// TIA Portal V20 export
FUNCTION_BLOCK "PR_FibroMainSeq_Soft2.0 1_workflow_a30ae2"   // FB43, LAD
{ S7_Optimized_Access := 'TRUE' }
// stored: MemoryReserve 100, SetENOAutomatically false
   VAR_INPUT
      iAllStationsSafe : Bool;
      iAllTaskOver : Bool;
      iAutoRunning : Bool;
      iFaultReset : Bool;
      iFibroAtStnPos : Bool;
      iIndexOver : Bool;
      iProcessActive : Bool;
      iReset_fault : Bool;
      iSstMode : Bool;
      iSstPB : Bool;
   END_VAR
   VAR_OUTPUT
      qError : Array[1..1] of Bool;
      qMessage_0 : Bool;
      qProcessActive : Bool;
   END_VAR
   VAR
      c10_ChkRecCond_T1 : Bool;
      c10_ChkRecCond_T2 : Bool;
      c10_ChkRecCond_T3 : Bool;
      c50_ChkPartPresentAtStn_T1 : Bool;
      c50_ChkPartPresentAtStn_T2 : Bool;
      StateNo : Int;
      s100_WtAllStnTaskOver : Bool;
      s100_WtAllStnTaskOver_T1 : Bool;
      s10_ChkRecCond : Bool;
      s10_ChkRecCond_T1 : Bool;
      s10_ChkRecCond_T2 : Bool;
      s10_ChkRecCond_T3 : Bool;
      s130_ChkAllStnSafe2 : Bool;
      s130_ChkAllStnSafe2_T1 : Bool;
      s140_WtIndexOver : Bool;
      s140_WtIndexOver_T1 : Bool;
      s1_WtResetRel : Bool;
      s1_WtResetRel_T1 : Bool;
      s20_WtManualIntv : Bool;
      s20_WtManualIntv_T1 : Bool;
      s30_WtFibroAtStnPos : Bool;
      s30_WtFibroAtStnPos_T1 : Bool;
      s40_ChkAllStnSafe : Bool;
      s40_ChkAllStnSafe_T1 : Bool;
      s50_ChkPartPresentAtStn : Bool;
      s50_ChkPartPresentAtStn_T1 : Bool;
      s50_ChkPartPresentAtStn_T2 : Bool;
      s60_WtPartPresentAtStn : Bool;
      s60_WtPartPresentAtStn_T1 : Bool;
      sAbnormalCondition : Bool;
      sPartPresentAtStation : Bool;
      sProcessActive : Bool;
      sSst : Bool;
      sSstPulse : Bool;
      sSstRise : Bool;
      sStWtResetRel : Bool;
      sStWtResetRel_T1 : Bool;
   END_VAR
   VAR_TEMP
      tOne : Bool;
   END_VAR
   VAR_TEMP   // added for the SCL form of the ladder/FBD networks
      _w1 : Bool;
      _w2 : Bool;
   END_VAR
BEGIN

REGION Network 1
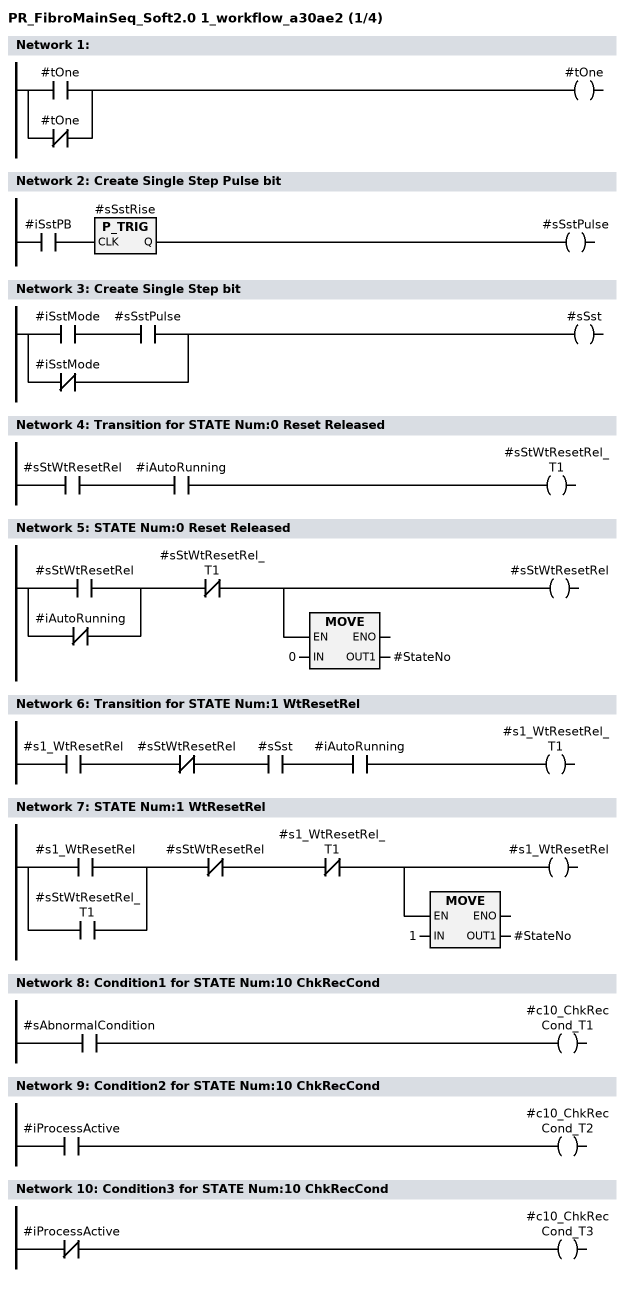
   RUNG wire#powerrail
      Contact( #tOne )
      wire#w1
      Coil( #tOne )
   END_RUNG
   RUNG wire#powerrail
      I_Contact( #tOne )
   END_RUNG wire#w1
   // the same network as SCL:
   #tOne := #tOne OR NOT #tOne;
END_REGION

REGION Network 2: Create Single Step Pulse bit
   RUNG wire#powerrail
      Contact( #iSstPB )
      P_Trig( #sSstRise )
      Coil( #sSstPulse )
   END_RUNG
   // the same network as SCL:
   #_w1 := #iSstPB AND NOT #sSstRise;   // rising edge
   #sSstRise := #iSstPB;
   #sSstPulse := #_w1;
END_REGION

REGION Network 3: Create Single Step bit
   RUNG wire#powerrail
      Contact( #iSstMode )
      Contact( #sSstPulse )
      wire#w1
      Coil( #sSst )
   END_RUNG
   RUNG wire#powerrail
      I_Contact( #iSstMode )
   END_RUNG wire#w1
   // the same network as SCL:
   #sSst := (#iSstMode AND #sSstPulse) OR NOT #iSstMode;
END_REGION

REGION Network 4: Transition for STATE Num:0 Reset Released
   RUNG wire#powerrail
      Contact( #sStWtResetRel )
      Contact( #iAutoRunning )
      Coil( #sStWtResetRel_T1 )
   END_RUNG
   // the same network as SCL:
   #sStWtResetRel_T1 := #sStWtResetRel AND #iAutoRunning;
END_REGION

REGION Network 5: STATE Num:0 Reset Released
   RUNG wire#powerrail
      Contact( #sStWtResetRel )
      wire#w1
      I_Contact( #sStWtResetRel_T1 )
      wire#w2
      Coil( #sStWtResetRel )
   END_RUNG
   RUNG wire#powerrail
      I_Contact( #iAutoRunning )
   END_RUNG wire#w1
   RUNG wire#w2
      { S7_GenerateENO := "TRUE" } Move(in := 0, out1 => #StateNo)
   END_RUNG
   // the same network as SCL:
   #sStWtResetRel := (#sStWtResetRel OR NOT #iAutoRunning) AND NOT #sStWtResetRel_T1;
   IF #sStWtResetRel THEN #StateNo := 0; END_IF;
END_REGION

REGION Network 6: Transition for STATE Num:1 WtResetRel
   RUNG wire#powerrail
      Contact( #s1_WtResetRel )
      I_Contact( #sStWtResetRel )
      Contact( #sSst )
      Contact( #iAutoRunning )
      Coil( #s1_WtResetRel_T1 )
   END_RUNG
   // the same network as SCL:
   #s1_WtResetRel_T1 := #s1_WtResetRel AND NOT #sStWtResetRel AND #sSst AND #iAutoRunning;
END_REGION

REGION Network 7: STATE Num:1 WtResetRel
   RUNG wire#powerrail
      Contact( #s1_WtResetRel )
      wire#w1
      I_Contact( #sStWtResetRel )
      I_Contact( #s1_WtResetRel_T1 )
      wire#w2
      Coil( #s1_WtResetRel )
   END_RUNG
   RUNG wire#powerrail
      Contact( #sStWtResetRel_T1 )
   END_RUNG wire#w1
   RUNG wire#w2
      { S7_GenerateENO := "TRUE" } Move(in := 1, out1 => #StateNo)
   END_RUNG
   // the same network as SCL:
   #s1_WtResetRel := (#s1_WtResetRel OR #sStWtResetRel_T1) AND NOT #sStWtResetRel AND NOT #s1_WtResetRel_T1;
   IF #s1_WtResetRel THEN #StateNo := 1; END_IF;
END_REGION

REGION Network 8: Condition1 for STATE Num:10 ChkRecCond
   RUNG wire#powerrail
      Contact( #sAbnormalCondition )
      Coil( #c10_ChkRecCond_T1 )
   END_RUNG
   // the same network as SCL:
   #c10_ChkRecCond_T1 := #sAbnormalCondition;
END_REGION

REGION Network 9: Condition2 for STATE Num:10 ChkRecCond
   RUNG wire#powerrail
      Contact( #iProcessActive )
      Coil( #c10_ChkRecCond_T2 )
   END_RUNG
   // the same network as SCL:
   #c10_ChkRecCond_T2 := #iProcessActive;
END_REGION

REGION Network 10: Condition3 for STATE Num:10 ChkRecCond
   RUNG wire#powerrail
      I_Contact( #iProcessActive )
      Coil( #c10_ChkRecCond_T3 )
   END_RUNG
   // the same network as SCL:
   #c10_ChkRecCond_T3 := NOT #iProcessActive;
END_REGION

REGION Network 11: Transition for STATE Num:10 ChkRecCond
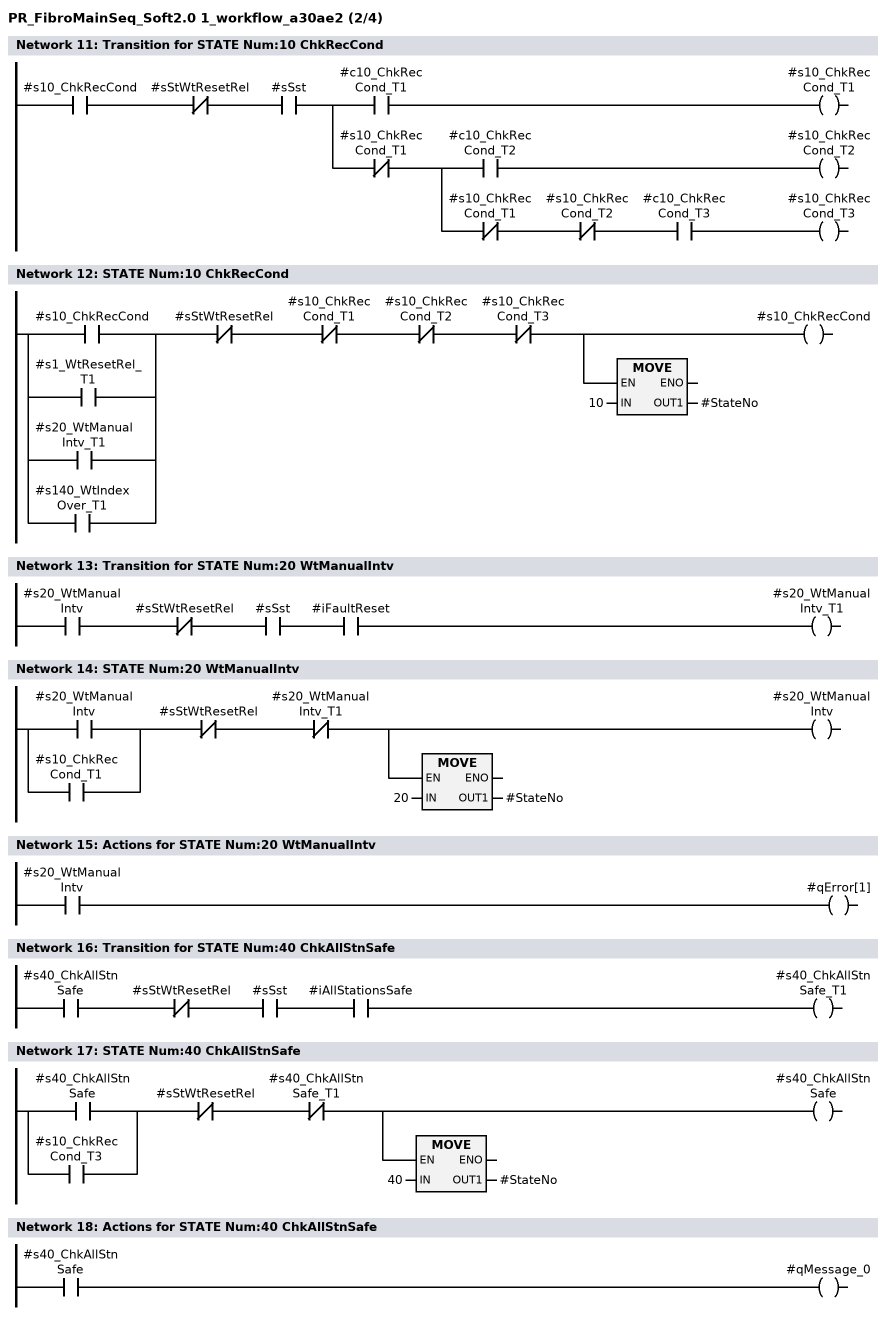
   RUNG wire#powerrail
      Contact( #s10_ChkRecCond )
      I_Contact( #sStWtResetRel )
      Contact( #sSst )
      wire#w1
      Contact( #c10_ChkRecCond_T1 )
      Coil( #s10_ChkRecCond_T1 )
   END_RUNG
   RUNG wire#w1
      I_Contact( #s10_ChkRecCond_T1 )
      wire#w2
      Contact( #c10_ChkRecCond_T2 )
      Coil( #s10_ChkRecCond_T2 )
   END_RUNG
   RUNG wire#w2
      I_Contact( #s10_ChkRecCond_T1 )
      I_Contact( #s10_ChkRecCond_T2 )
      Contact( #c10_ChkRecCond_T3 )
      Coil( #s10_ChkRecCond_T3 )
   END_RUNG
   // the same network as SCL:
   #_w1 := #s10_ChkRecCond AND NOT #sStWtResetRel AND #sSst;
   #s10_ChkRecCond_T1 := #_w1 AND #c10_ChkRecCond_T1;
   #_w2 := #_w1 AND NOT #s10_ChkRecCond_T1;
   #s10_ChkRecCond_T2 := #_w2 AND #c10_ChkRecCond_T2;
   #s10_ChkRecCond_T3 := #_w2 AND NOT #s10_ChkRecCond_T1 AND NOT #s10_ChkRecCond_T2 AND #c10_ChkRecCond_T3;
END_REGION

REGION Network 12: STATE Num:10 ChkRecCond
   RUNG wire#powerrail
      Contact( #s10_ChkRecCond )
      wire#w1
      I_Contact( #sStWtResetRel )
      I_Contact( #s10_ChkRecCond_T1 )
      I_Contact( #s10_ChkRecCond_T2 )
      I_Contact( #s10_ChkRecCond_T3 )
      wire#w2
      Coil( #s10_ChkRecCond )
   END_RUNG
   RUNG wire#powerrail
      Contact( #s1_WtResetRel_T1 )
   END_RUNG wire#w1
   RUNG wire#powerrail
      Contact( #s20_WtManualIntv_T1 )
   END_RUNG wire#w1
   RUNG wire#powerrail
      Contact( #s140_WtIndexOver_T1 )
   END_RUNG wire#w1
   RUNG wire#w2
      { S7_GenerateENO := "TRUE" } Move(in := 10, out1 => #StateNo)
   END_RUNG
   // the same network as SCL:
   #s10_ChkRecCond := (#s10_ChkRecCond OR #s1_WtResetRel_T1 OR #s20_WtManualIntv_T1 OR #s140_WtIndexOver_T1) AND NOT #sStWtResetRel AND NOT #s10_ChkRecCond_T1 AND NOT #s10_ChkRecCond_T2 AND NOT #s10_ChkRecCond_T3;
   IF #s10_ChkRecCond THEN #StateNo := 10; END_IF;
END_REGION

REGION Network 13: Transition for STATE Num:20 WtManualIntv
   RUNG wire#powerrail
      Contact( #s20_WtManualIntv )
      I_Contact( #sStWtResetRel )
      Contact( #sSst )
      Contact( #iFaultReset )
      Coil( #s20_WtManualIntv_T1 )
   END_RUNG
   // the same network as SCL:
   #s20_WtManualIntv_T1 := #s20_WtManualIntv AND NOT #sStWtResetRel AND #sSst AND #iFaultReset;
END_REGION

REGION Network 14: STATE Num:20 WtManualIntv
   RUNG wire#powerrail
      Contact( #s20_WtManualIntv )
      wire#w1
      I_Contact( #sStWtResetRel )
      I_Contact( #s20_WtManualIntv_T1 )
      wire#w2
      Coil( #s20_WtManualIntv )
   END_RUNG
   RUNG wire#powerrail
      Contact( #s10_ChkRecCond_T1 )
   END_RUNG wire#w1
   RUNG wire#w2
      { S7_GenerateENO := "TRUE" } Move(in := 20, out1 => #StateNo)
   END_RUNG
   // the same network as SCL:
   #s20_WtManualIntv := (#s20_WtManualIntv OR #s10_ChkRecCond_T1) AND NOT #sStWtResetRel AND NOT #s20_WtManualIntv_T1;
   IF #s20_WtManualIntv THEN #StateNo := 20; END_IF;
END_REGION

REGION Network 15: Actions for STATE Num:20 WtManualIntv
   RUNG wire#powerrail
      Contact( #s20_WtManualIntv )
      Coil( #qError[1] )
   END_RUNG
   // the same network as SCL:
   #qError[1] := #s20_WtManualIntv;
END_REGION

REGION Network 16: Transition for STATE Num:40 ChkAllStnSafe
   RUNG wire#powerrail
      Contact( #s40_ChkAllStnSafe )
      I_Contact( #sStWtResetRel )
      Contact( #sSst )
      Contact( #iAllStationsSafe )
      Coil( #s40_ChkAllStnSafe_T1 )
   END_RUNG
   // the same network as SCL:
   #s40_ChkAllStnSafe_T1 := #s40_ChkAllStnSafe AND NOT #sStWtResetRel AND #sSst AND #iAllStationsSafe;
END_REGION

REGION Network 17: STATE Num:40 ChkAllStnSafe
   RUNG wire#powerrail
      Contact( #s40_ChkAllStnSafe )
      wire#w1
      I_Contact( #sStWtResetRel )
      I_Contact( #s40_ChkAllStnSafe_T1 )
      wire#w2
      Coil( #s40_ChkAllStnSafe )
   END_RUNG
   RUNG wire#powerrail
      Contact( #s10_ChkRecCond_T3 )
   END_RUNG wire#w1
   RUNG wire#w2
      { S7_GenerateENO := "TRUE" } Move(in := 40, out1 => #StateNo)
   END_RUNG
   // the same network as SCL:
   #s40_ChkAllStnSafe := (#s40_ChkAllStnSafe OR #s10_ChkRecCond_T3) AND NOT #sStWtResetRel AND NOT #s40_ChkAllStnSafe_T1;
   IF #s40_ChkAllStnSafe THEN #StateNo := 40; END_IF;
END_REGION

REGION Network 18: Actions for STATE Num:40 ChkAllStnSafe
   RUNG wire#powerrail
      Contact( #s40_ChkAllStnSafe )
      Coil( #qMessage_0 )
   END_RUNG
   // the same network as SCL:
   #qMessage_0 := #s40_ChkAllStnSafe;
END_REGION

REGION Network 19: Transition for STATE Num:30 WtFibroAtStnPos
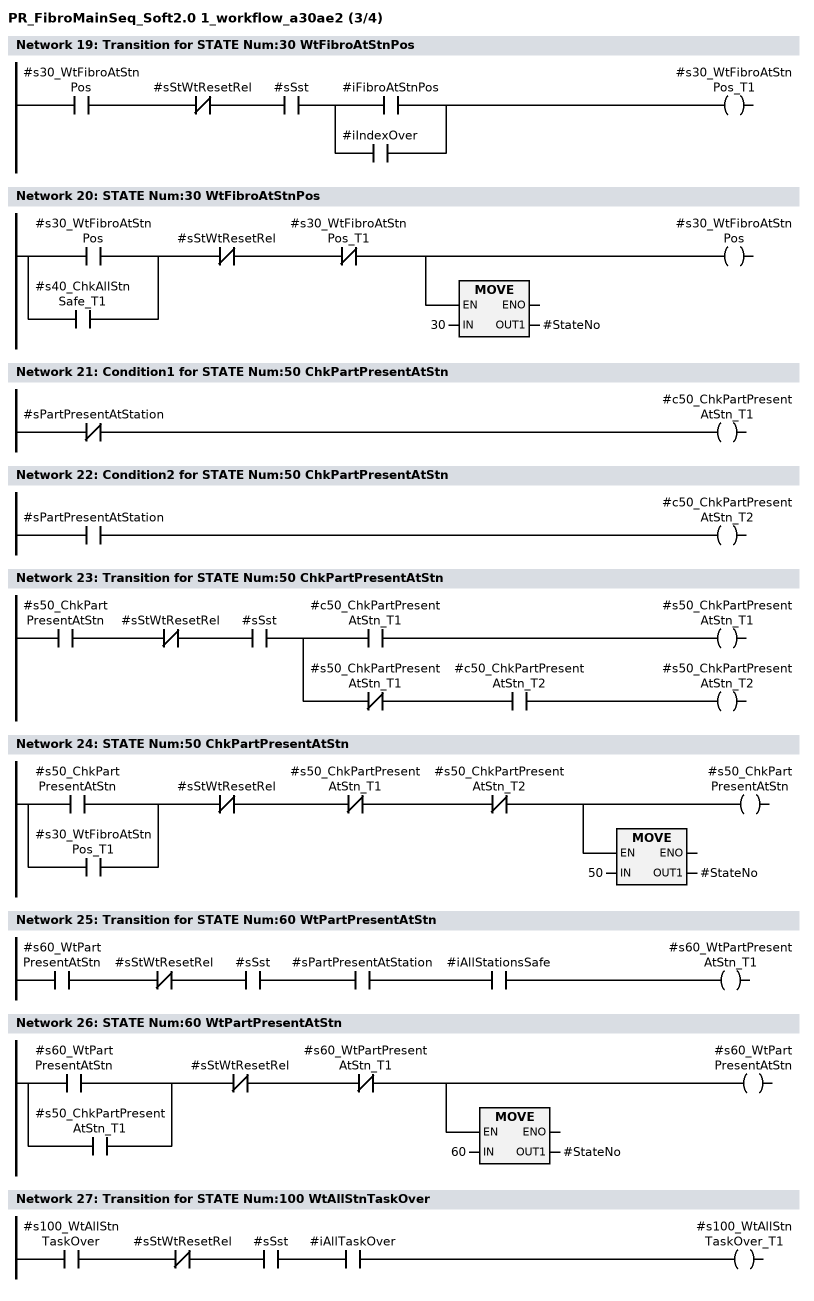
   RUNG wire#powerrail
      Contact( #s30_WtFibroAtStnPos )
      I_Contact( #sStWtResetRel )
      Contact( #sSst )
      wire#w1
      Contact( #iFibroAtStnPos )
      wire#w2
      Coil( #s30_WtFibroAtStnPos_T1 )
   END_RUNG
   RUNG wire#w1
      Contact( #iIndexOver )
   END_RUNG wire#w2
   // the same network as SCL:
   #s30_WtFibroAtStnPos_T1 := #s30_WtFibroAtStnPos AND NOT #sStWtResetRel AND #sSst AND (#iFibroAtStnPos OR #iIndexOver);
END_REGION

REGION Network 20: STATE Num:30 WtFibroAtStnPos
   RUNG wire#powerrail
      Contact( #s30_WtFibroAtStnPos )
      wire#w1
      I_Contact( #sStWtResetRel )
      I_Contact( #s30_WtFibroAtStnPos_T1 )
      wire#w2
      Coil( #s30_WtFibroAtStnPos )
   END_RUNG
   RUNG wire#powerrail
      Contact( #s40_ChkAllStnSafe_T1 )
   END_RUNG wire#w1
   RUNG wire#w2
      { S7_GenerateENO := "TRUE" } Move(in := 30, out1 => #StateNo)
   END_RUNG
   // the same network as SCL:
   #s30_WtFibroAtStnPos := (#s30_WtFibroAtStnPos OR #s40_ChkAllStnSafe_T1) AND NOT #sStWtResetRel AND NOT #s30_WtFibroAtStnPos_T1;
   IF #s30_WtFibroAtStnPos THEN #StateNo := 30; END_IF;
END_REGION

REGION Network 21: Condition1 for STATE Num:50 ChkPartPresentAtStn
   RUNG wire#powerrail
      I_Contact( #sPartPresentAtStation )
      Coil( #c50_ChkPartPresentAtStn_T1 )
   END_RUNG
   // the same network as SCL:
   #c50_ChkPartPresentAtStn_T1 := NOT #sPartPresentAtStation;
END_REGION

REGION Network 22: Condition2 for STATE Num:50 ChkPartPresentAtStn
   RUNG wire#powerrail
      Contact( #sPartPresentAtStation )
      Coil( #c50_ChkPartPresentAtStn_T2 )
   END_RUNG
   // the same network as SCL:
   #c50_ChkPartPresentAtStn_T2 := #sPartPresentAtStation;
END_REGION

REGION Network 23: Transition for STATE Num:50 ChkPartPresentAtStn
   RUNG wire#powerrail
      Contact( #s50_ChkPartPresentAtStn )
      I_Contact( #sStWtResetRel )
      Contact( #sSst )
      wire#w1
      Contact( #c50_ChkPartPresentAtStn_T1 )
      Coil( #s50_ChkPartPresentAtStn_T1 )
   END_RUNG
   RUNG wire#w1
      I_Contact( #s50_ChkPartPresentAtStn_T1 )
      Contact( #c50_ChkPartPresentAtStn_T2 )
      Coil( #s50_ChkPartPresentAtStn_T2 )
   END_RUNG
   // the same network as SCL:
   #_w1 := #s50_ChkPartPresentAtStn AND NOT #sStWtResetRel AND #sSst;
   #s50_ChkPartPresentAtStn_T1 := #_w1 AND #c50_ChkPartPresentAtStn_T1;
   #s50_ChkPartPresentAtStn_T2 := #_w1 AND NOT #s50_ChkPartPresentAtStn_T1 AND #c50_ChkPartPresentAtStn_T2;
END_REGION

REGION Network 24: STATE Num:50 ChkPartPresentAtStn
   RUNG wire#powerrail
      Contact( #s50_ChkPartPresentAtStn )
      wire#w1
      I_Contact( #sStWtResetRel )
      I_Contact( #s50_ChkPartPresentAtStn_T1 )
      I_Contact( #s50_ChkPartPresentAtStn_T2 )
      wire#w2
      Coil( #s50_ChkPartPresentAtStn )
   END_RUNG
   RUNG wire#powerrail
      Contact( #s30_WtFibroAtStnPos_T1 )
   END_RUNG wire#w1
   RUNG wire#w2
      { S7_GenerateENO := "TRUE" } Move(in := 50, out1 => #StateNo)
   END_RUNG
   // the same network as SCL:
   #s50_ChkPartPresentAtStn := (#s50_ChkPartPresentAtStn OR #s30_WtFibroAtStnPos_T1) AND NOT #sStWtResetRel AND NOT #s50_ChkPartPresentAtStn_T1 AND NOT #s50_ChkPartPresentAtStn_T2;
   IF #s50_ChkPartPresentAtStn THEN #StateNo := 50; END_IF;
END_REGION

REGION Network 25: Transition for STATE Num:60 WtPartPresentAtStn
   RUNG wire#powerrail
      Contact( #s60_WtPartPresentAtStn )
      I_Contact( #sStWtResetRel )
      Contact( #sSst )
      Contact( #sPartPresentAtStation )
      Contact( #iAllStationsSafe )
      Coil( #s60_WtPartPresentAtStn_T1 )
   END_RUNG
   // the same network as SCL:
   #s60_WtPartPresentAtStn_T1 := #s60_WtPartPresentAtStn AND NOT #sStWtResetRel AND #sSst AND #sPartPresentAtStation AND #iAllStationsSafe;
END_REGION

REGION Network 26: STATE Num:60 WtPartPresentAtStn
   RUNG wire#powerrail
      Contact( #s60_WtPartPresentAtStn )
      wire#w1
      I_Contact( #sStWtResetRel )
      I_Contact( #s60_WtPartPresentAtStn_T1 )
      wire#w2
      Coil( #s60_WtPartPresentAtStn )
   END_RUNG
   RUNG wire#powerrail
      Contact( #s50_ChkPartPresentAtStn_T1 )
   END_RUNG wire#w1
   RUNG wire#w2
      { S7_GenerateENO := "TRUE" } Move(in := 60, out1 => #StateNo)
   END_RUNG
   // the same network as SCL:
   #s60_WtPartPresentAtStn := (#s60_WtPartPresentAtStn OR #s50_ChkPartPresentAtStn_T1) AND NOT #sStWtResetRel AND NOT #s60_WtPartPresentAtStn_T1;
   IF #s60_WtPartPresentAtStn THEN #StateNo := 60; END_IF;
END_REGION

REGION Network 27: Transition for STATE Num:100 WtAllStnTaskOver
   RUNG wire#powerrail
      Contact( #s100_WtAllStnTaskOver )
      I_Contact( #sStWtResetRel )
      Contact( #sSst )
      Contact( #iAllTaskOver )
      Coil( #s100_WtAllStnTaskOver_T1 )
   END_RUNG
   // the same network as SCL:
   #s100_WtAllStnTaskOver_T1 := #s100_WtAllStnTaskOver AND NOT #sStWtResetRel AND #sSst AND #iAllTaskOver;
END_REGION

REGION Network 28: STATE Num:100 WtAllStnTaskOver
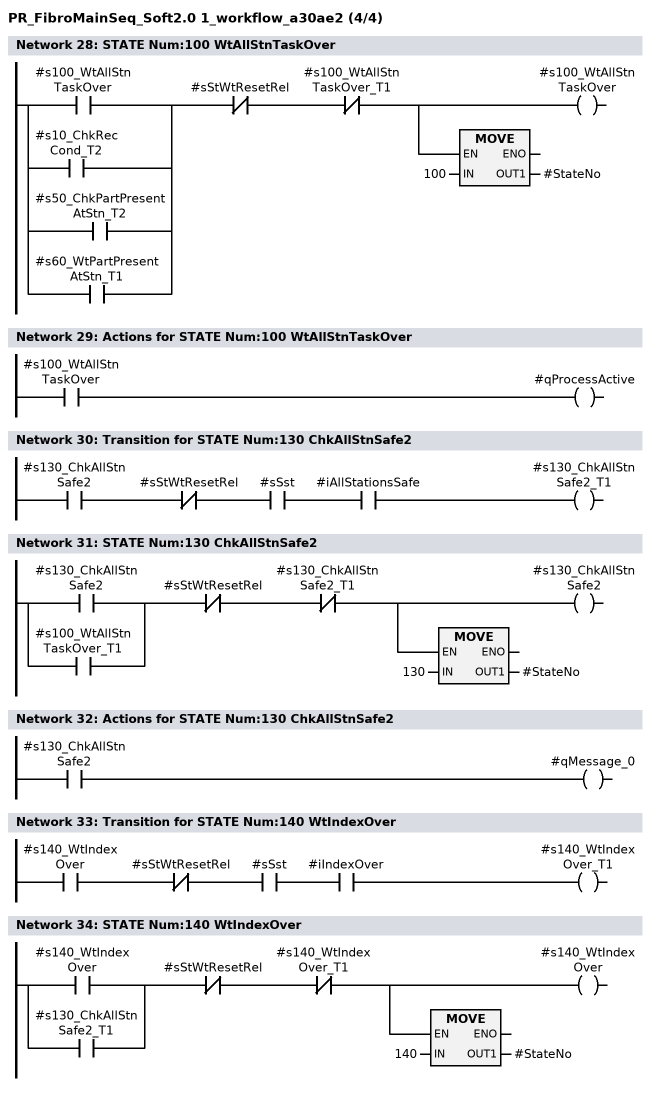
   RUNG wire#powerrail
      Contact( #s100_WtAllStnTaskOver )
      wire#w1
      I_Contact( #sStWtResetRel )
      I_Contact( #s100_WtAllStnTaskOver_T1 )
      wire#w2
      Coil( #s100_WtAllStnTaskOver )
   END_RUNG
   RUNG wire#powerrail
      Contact( #s10_ChkRecCond_T2 )
   END_RUNG wire#w1
   RUNG wire#powerrail
      Contact( #s50_ChkPartPresentAtStn_T2 )
   END_RUNG wire#w1
   RUNG wire#powerrail
      Contact( #s60_WtPartPresentAtStn_T1 )
   END_RUNG wire#w1
   RUNG wire#w2
      { S7_GenerateENO := "TRUE" } Move(in := 100, out1 => #StateNo)
   END_RUNG
   // the same network as SCL:
   #s100_WtAllStnTaskOver := (#s100_WtAllStnTaskOver OR #s10_ChkRecCond_T2 OR #s50_ChkPartPresentAtStn_T2 OR #s60_WtPartPresentAtStn_T1) AND NOT #sStWtResetRel AND NOT #s100_WtAllStnTaskOver_T1;
   IF #s100_WtAllStnTaskOver THEN #StateNo := 100; END_IF;
END_REGION

REGION Network 29: Actions for STATE Num:100 WtAllStnTaskOver
   RUNG wire#powerrail
      Contact( #s100_WtAllStnTaskOver )
      Coil( #qProcessActive )
   END_RUNG
   // the same network as SCL:
   #qProcessActive := #s100_WtAllStnTaskOver;
END_REGION

REGION Network 30: Transition for STATE Num:130 ChkAllStnSafe2
   RUNG wire#powerrail
      Contact( #s130_ChkAllStnSafe2 )
      I_Contact( #sStWtResetRel )
      Contact( #sSst )
      Contact( #iAllStationsSafe )
      Coil( #s130_ChkAllStnSafe2_T1 )
   END_RUNG
   // the same network as SCL:
   #s130_ChkAllStnSafe2_T1 := #s130_ChkAllStnSafe2 AND NOT #sStWtResetRel AND #sSst AND #iAllStationsSafe;
END_REGION

REGION Network 31: STATE Num:130 ChkAllStnSafe2
   RUNG wire#powerrail
      Contact( #s130_ChkAllStnSafe2 )
      wire#w1
      I_Contact( #sStWtResetRel )
      I_Contact( #s130_ChkAllStnSafe2_T1 )
      wire#w2
      Coil( #s130_ChkAllStnSafe2 )
   END_RUNG
   RUNG wire#powerrail
      Contact( #s100_WtAllStnTaskOver_T1 )
   END_RUNG wire#w1
   RUNG wire#w2
      { S7_GenerateENO := "TRUE" } Move(in := 130, out1 => #StateNo)
   END_RUNG
   // the same network as SCL:
   #s130_ChkAllStnSafe2 := (#s130_ChkAllStnSafe2 OR #s100_WtAllStnTaskOver_T1) AND NOT #sStWtResetRel AND NOT #s130_ChkAllStnSafe2_T1;
   IF #s130_ChkAllStnSafe2 THEN #StateNo := 130; END_IF;
END_REGION

REGION Network 32: Actions for STATE Num:130 ChkAllStnSafe2
   RUNG wire#powerrail
      Contact( #s130_ChkAllStnSafe2 )
      Coil( #qMessage_0 )
   END_RUNG
   // the same network as SCL:
   #qMessage_0 := #s130_ChkAllStnSafe2;
END_REGION

REGION Network 33: Transition for STATE Num:140 WtIndexOver
   RUNG wire#powerrail
      Contact( #s140_WtIndexOver )
      I_Contact( #sStWtResetRel )
      Contact( #sSst )
      Contact( #iIndexOver )
      Coil( #s140_WtIndexOver_T1 )
   END_RUNG
   // the same network as SCL:
   #s140_WtIndexOver_T1 := #s140_WtIndexOver AND NOT #sStWtResetRel AND #sSst AND #iIndexOver;
END_REGION

REGION Network 34: STATE Num:140 WtIndexOver
   RUNG wire#powerrail
      Contact( #s140_WtIndexOver )
      wire#w1
      I_Contact( #sStWtResetRel )
      I_Contact( #s140_WtIndexOver_T1 )
      wire#w2
      Coil( #s140_WtIndexOver )
   END_RUNG
   RUNG wire#powerrail
      Contact( #s130_ChkAllStnSafe2_T1 )
   END_RUNG wire#w1
   RUNG wire#w2
      { S7_GenerateENO := "TRUE" } Move(in := 140, out1 => #StateNo)
   END_RUNG
   // the same network as SCL:
   #s140_WtIndexOver := (#s140_WtIndexOver OR #s130_ChkAllStnSafe2_T1) AND NOT #sStWtResetRel AND NOT #s140_WtIndexOver_T1;
   IF #s140_WtIndexOver THEN #StateNo := 140; END_IF;
END_REGION
END_FUNCTION_BLOCK
